// TIA Portal V20 export
ORGANIZATION_BLOCK "T5_Ciclo"   // OB128, LAD, ProgramCycle
TITLE = T5_Ciclo
{ S7_Optimized_Access := 'TRUE' }
AUTHOR : IA
FAMILY : PRUEBA
VERSION : 0.1
// Tanda 1b: llama a todas las pruebas
// stored: AutoNumber false, IsIECCheckEnabled false, SetENOAutomatically false
   VAR_INPUT
      Initial_Call : Bool;
      Remanence : Bool;
   END_VAR
BEGIN

REGION Network 1: T5_Base
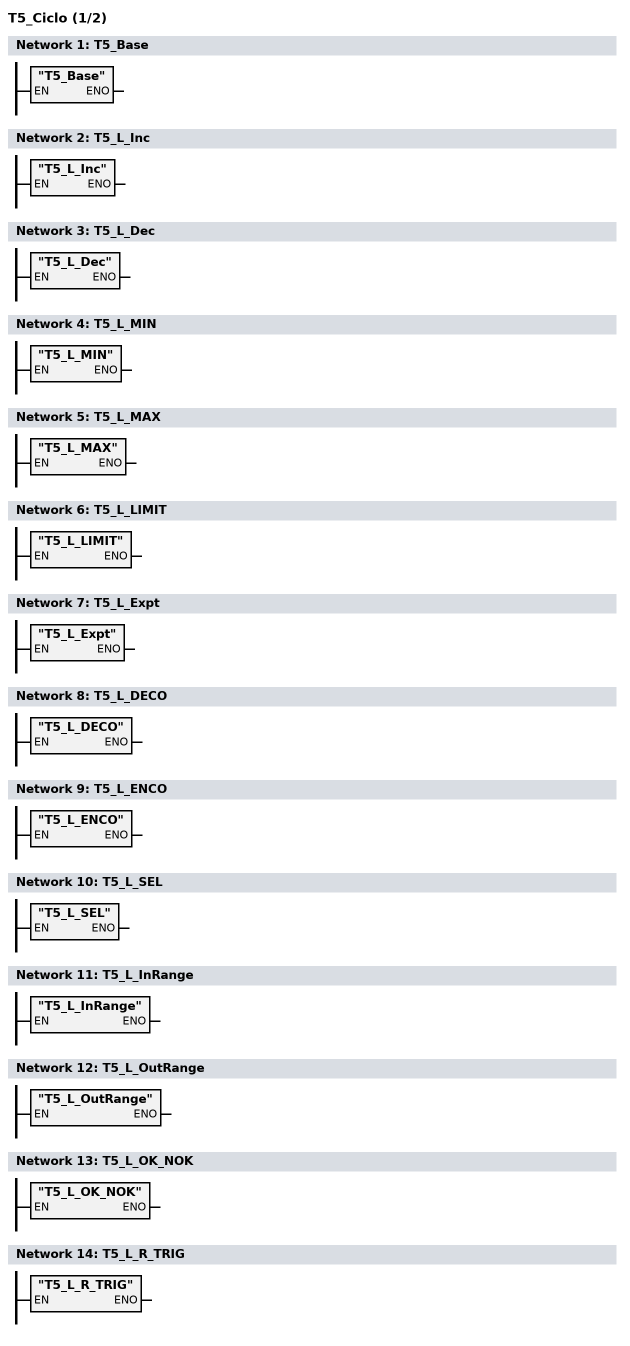
   RUNG wire#powerrail
      "T5_Base"()
   END_RUNG
   // the same network as SCL:
   "T5_Base"();
END_REGION

REGION Network 2: T5_L_Inc
   RUNG wire#powerrail
      "T5_L_Inc"()
   END_RUNG
   // the same network as SCL:
   "T5_L_Inc"();
END_REGION

REGION Network 3: T5_L_Dec
   RUNG wire#powerrail
      "T5_L_Dec"()
   END_RUNG
   // the same network as SCL:
   "T5_L_Dec"();
END_REGION

REGION Network 4: T5_L_MIN
   RUNG wire#powerrail
      "T5_L_MIN"()
   END_RUNG
   // the same network as SCL:
   "T5_L_MIN"();
END_REGION

REGION Network 5: T5_L_MAX
   RUNG wire#powerrail
      "T5_L_MAX"()
   END_RUNG
   // the same network as SCL:
   "T5_L_MAX"();
END_REGION

REGION Network 6: T5_L_LIMIT
   RUNG wire#powerrail
      "T5_L_LIMIT"()
   END_RUNG
   // the same network as SCL:
   "T5_L_LIMIT"();
END_REGION

REGION Network 7: T5_L_Expt
   RUNG wire#powerrail
      "T5_L_Expt"()
   END_RUNG
   // the same network as SCL:
   "T5_L_Expt"();
END_REGION

REGION Network 8: T5_L_DECO
   RUNG wire#powerrail
      "T5_L_DECO"()
   END_RUNG
   // the same network as SCL:
   "T5_L_DECO"();
END_REGION

REGION Network 9: T5_L_ENCO
   RUNG wire#powerrail
      "T5_L_ENCO"()
   END_RUNG
   // the same network as SCL:
   "T5_L_ENCO"();
END_REGION

REGION Network 10: T5_L_SEL
   RUNG wire#powerrail
      "T5_L_SEL"()
   END_RUNG
   // the same network as SCL:
   "T5_L_SEL"();
END_REGION

REGION Network 11: T5_L_InRange
   RUNG wire#powerrail
      "T5_L_InRange"()
   END_RUNG
   // the same network as SCL:
   "T5_L_InRange"();
END_REGION

REGION Network 12: T5_L_OutRange
   RUNG wire#powerrail
      "T5_L_OutRange"()
   END_RUNG
   // the same network as SCL:
   "T5_L_OutRange"();
END_REGION

REGION Network 13: T5_L_OK_NOK
   RUNG wire#powerrail
      "T5_L_OK_NOK"()
   END_RUNG
   // the same network as SCL:
   "T5_L_OK_NOK"();
END_REGION

REGION Network 14: T5_L_R_TRIG
   RUNG wire#powerrail
      "T5_L_R_TRIG"()
   END_RUNG
   // the same network as SCL:
   "T5_L_R_TRIG"();
END_REGION

REGION Network 15: T5_L_F_TRIG
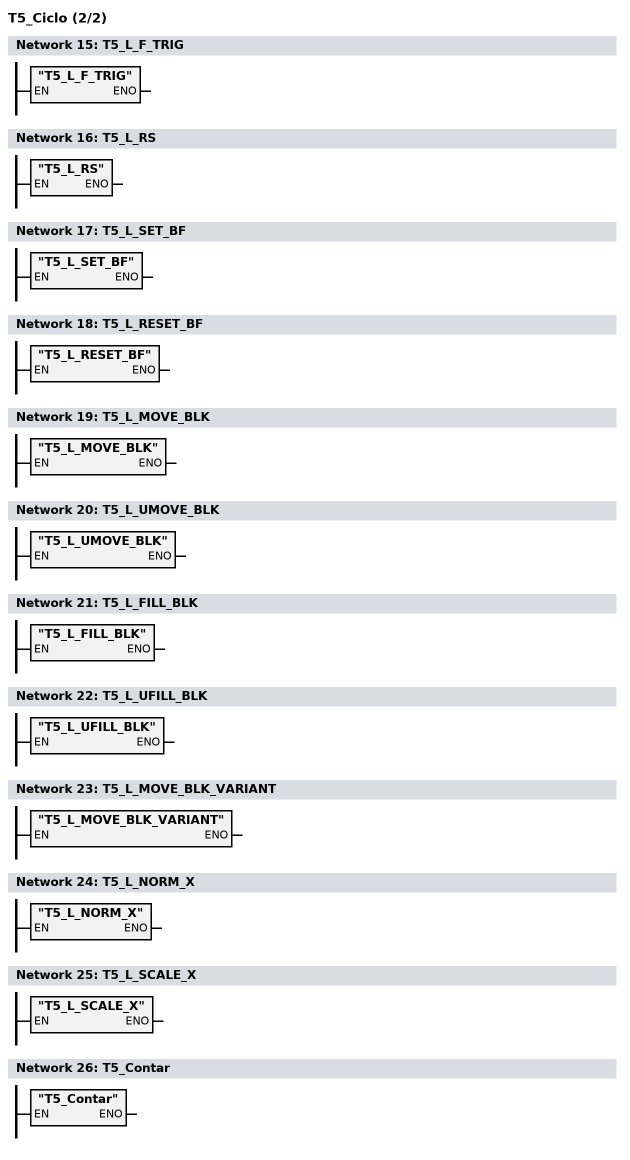
   RUNG wire#powerrail
      "T5_L_F_TRIG"()
   END_RUNG
   // the same network as SCL:
   "T5_L_F_TRIG"();
END_REGION

REGION Network 16: T5_L_RS
   RUNG wire#powerrail
      "T5_L_RS"()
   END_RUNG
   // the same network as SCL:
   "T5_L_RS"();
END_REGION

REGION Network 17: T5_L_SET_BF
   RUNG wire#powerrail
      "T5_L_SET_BF"()
   END_RUNG
   // the same network as SCL:
   "T5_L_SET_BF"();
END_REGION

REGION Network 18: T5_L_RESET_BF
   RUNG wire#powerrail
      "T5_L_RESET_BF"()
   END_RUNG
   // the same network as SCL:
   "T5_L_RESET_BF"();
END_REGION

REGION Network 19: T5_L_MOVE_BLK
   RUNG wire#powerrail
      "T5_L_MOVE_BLK"()
   END_RUNG
   // the same network as SCL:
   "T5_L_MOVE_BLK"();
END_REGION

REGION Network 20: T5_L_UMOVE_BLK
   RUNG wire#powerrail
      "T5_L_UMOVE_BLK"()
   END_RUNG
   // the same network as SCL:
   "T5_L_UMOVE_BLK"();
END_REGION

REGION Network 21: T5_L_FILL_BLK
   RUNG wire#powerrail
      "T5_L_FILL_BLK"()
   END_RUNG
   // the same network as SCL:
   "T5_L_FILL_BLK"();
END_REGION

REGION Network 22: T5_L_UFILL_BLK
   RUNG wire#powerrail
      "T5_L_UFILL_BLK"()
   END_RUNG
   // the same network as SCL:
   "T5_L_UFILL_BLK"();
END_REGION

REGION Network 23: T5_L_MOVE_BLK_VARIANT
   RUNG wire#powerrail
      "T5_L_MOVE_BLK_VARIANT"()
   END_RUNG
   // the same network as SCL:
   "T5_L_MOVE_BLK_VARIANT"();
END_REGION

REGION Network 24: T5_L_NORM_X
   RUNG wire#powerrail
      "T5_L_NORM_X"()
   END_RUNG
   // the same network as SCL:
   "T5_L_NORM_X"();
END_REGION

REGION Network 25: T5_L_SCALE_X
   RUNG wire#powerrail
      "T5_L_SCALE_X"()
   END_RUNG
   // the same network as SCL:
   "T5_L_SCALE_X"();
END_REGION

REGION Network 26: T5_Contar
   RUNG wire#powerrail
      "T5_Contar"()
   END_RUNG
   // the same network as SCL:
   "T5_Contar"();
END_REGION
END_ORGANIZATION_BLOCK
